// TwinCAT 3 PLC project Conveyor
// ProgramVersion: 3.1.4026.27
// libraries:
//   Tc2_Standard, * (Beckhoff Automation GmbH)
//   Tc2_System, * (Beckhoff Automation GmbH)
//   Tc3_Module, * (Beckhoff Automation GmbH)
// project tree:
//   GVLs/ GVL_IO.TcGVL
//   / PlcTask.TcTTO
//   POUs/ E_ConveyorMode.TcDUT, E_ConveyorState.TcDUT, E_FaultCode.TcDUT, FB_Conveyor.TcPOU, MAIN.TcPOU
// real-time tasks:
//   TASK PlcTask: cycle T#10ms, priority 20, ADS port 350

CONFIGURATION Conveyor
    RESOURCE PLC ON TwinCAT3
        TASK PlcTask(INTERVAL := T#10ms, PRIORITY := 20);
        PROGRAM MAIN WITH PlcTask : MAIN;
    END_RESOURCE
END_CONFIGURATION

// ---- POUs/E_ConveyorMode.TcDUT
{attribute 'qualified_only'}
{attribute 'strict'}
TYPE E_ConveyorMode  :
(
	AUTO,
	MANUAL
);
END_TYPE

// ---- POUs/E_ConveyorState.TcDUT
{attribute 'qualified_only'}
{attribute 'strict'}
TYPE E_ConveyorState :
(
	IDLE,
    RUNNING,
	WAIT_EXIT,
    FAULT
);
END_TYPE

// ---- POUs/E_FaultCode.TcDUT
{attribute 'qualified_only'}
{attribute 'strict'}
TYPE E_FaultCode :
(
	FC_NONE,
	FC_EMERGENCY_STOP,
	FC_EXIT_TIMEOUT
);
END_TYPE

// ---- GVLs/GVL_IO.TcGVL
{attribute 'qualified_only'}
VAR_GLOBAL
	//Input
	StartButton		:	BOOL;
	StopButton		:	BOOL;
	EmergencyStop	:	BOOL;
	Reset			:	BOOL;
	
	SensorEntry		:	BOOL;
	SensorExit		:	BOOL;
	AutoMode		:	BOOL;
	
	
	//Output
	Motor			:	BOOL;
	MotorStopped 	: 	BOOL;
	GreenLamp 		:	BOOL;
	RedLamp 		:	BOOL;
	
	FaultLamp		:	BOOL;
	
	FaultCode 		: 	E_FaultCode;
	
	FaultText : STRING(50) := 'NO FAULT';
	ModeText  : STRING(50) ;
	
	
	Mode : E_ConveyorMode := E_ConveyorMode.AUTO;
	
	
	
	
END_VAR

// ---- POUs/MAIN.TcPOU
PROGRAM MAIN
VAR
	Conveyor		:	FB_Conveyor;
	StartTrigger 	: 	R_TRIG;
	StopTrigger		:	R_TRIG;
	EmergencyOn		:	R_TRIG;
	Reset			:	R_TRIG; 
	
	
	
	
END_VAR

Conveyor(
    Start := GVL_IO.StartButton,
    Stop := GVL_IO.StopButton,
    EmergencyStop := GVL_IO.EmergencyStop,
    Reset := GVL_IO.Reset,
	AutoMode := GVL_IO.AutoMode,
	Mode := GVL_IO.Mode
);

GVL_IO.Motor := Conveyor.Motor;
GVL_IO.MotorStopped := NOT Conveyor.Motor;
GVL_IO.GreenLamp := Conveyor.GreenLamp;
GVL_IO.RedLamp := Conveyor.RedLamp;
GVL_IO.FaultLamp := Conveyor.FaultLamp;
GVL_IO.FaultCode := Conveyor.FaultCode;

GVL_IO.FaultCode := Conveyor.FaultCode;

IF GVL_IO.Mode = E_ConveyorMode.AUTO THEN
	StartTrigger(CLK := GVL_IO.StartButton);
END_IF

StopTrigger(CLK := GVL_IO.StopButton);
EmergencyOn(CLK:= GVL_IO.EmergencyStop);
Reset(CLK:=GVL_IO.Reset);


IF StartTrigger.Q THEN
    GVL_IO.StartButton := FALSE;
END_IF;
IF StopTrigger.Q THEN
	GVL_IO.StopButton := FALSE;
END_IF
IF EmergencyOn.Q THEN
	GVL_IO.EmergencyStop := FALSE;
END_IF
IF Reset.Q THEN
	GVL_IO.Reset := FALSE;
END_IF


CASE GVL_IO.FaultCode OF
    E_FaultCode.FC_NONE:
        GVL_IO.FaultText := 'NO FAULT';

    E_FaultCode.FC_EMERGENCY_STOP:
        GVL_IO.FaultText := 'EMERGENCY STOP';

    E_FaultCode.FC_EXIT_TIMEOUT:
        GVL_IO.FaultText := 'EXIT SENSOR TIMEOUT';
END_CASE

IF GVL_IO.AutoMode THEN
    GVL_IO.Mode := E_ConveyorMode.AUTO;
ELSE
    GVL_IO.Mode := E_ConveyorMode.MANUAL;
END_IF

IF GVL_IO.Mode = E_ConveyorMode.AUTO THEN
	GVL_IO.ModeText := 'AUTO';
ELSIF GVL_IO.Mode = E_ConveyorMode.MANUAL THEN
	GVL_IO.ModeText := 'MANUAL'; 
END_IF

END_PROGRAM

// ---- POUs/FB_Conveyor.TcPOU
FUNCTION_BLOCK FB_Conveyor
VAR_INPUT
	
	Start			:	BOOL;
	Stop			:	BOOL;
	EmergencyStop	:	BOOL;
	Reset			:	BOOL;
	
	AutoMode      	:	BOOL;
	SensorEntry   	: 	BOOL;
    SensorExit    	: 	BOOL;
	
	Mode	:	E_ConveyorMode;
	
END_VAR
VAR_OUTPUT
	
	Motor 		: BOOL;
	GreenLamp 	: BOOL;
	RedLamp 	: BOOL;
	FaultLamp	: BOOL;
	
	FaultCode : E_FaultCode := E_FaultCode.FC_NONE;
	
	
	
END_VAR
VAR
	
   
   
	
	State 	: 	E_ConveyorState ;
	
	
	ModeChanged 	: BOOL;
    PreviousMode 	: E_ConveyorMode;

  
	
	TimerPart		:	TON;
	ExitTrigger		:	R_TRIG;
	EntryTrigger 	: 	R_TRIG;
	Counter 		: 	UDINT := 0;
	
	InterlockOK 	: 	BOOL;
	
	
	
	
	
END_VAR

TimerPart(
    	IN := (Mode = E_ConveyorMode.AUTO)
          	AND 
				(State = E_ConveyorState.WAIT_EXIT),
    	PT := T#10S
	);
ExitTrigger(CLK := SensorExit);	
EntryTrigger(CLK := SensorEntry);
ModeChanged := Mode <> PreviousMode;

IF NOT HandleFaults() THEN
    IF NOT HandleModeChange() THEN
        IF Mode = E_ConveyorMode.AUTO THEN
            RunAuto();

        ELSIF Mode = E_ConveyorMode.MANUAL THEN
            RunManual();
        END_IF
    END_IF
END_IF

UpdateOutputs();

METHOD HandleFaults : BOOL
VAR_INPUT
END_VAR

VAR
END_VAR
HandleFaults := FALSE;

IF EmergencyStop THEN
    State := E_ConveyorState.FAULT;
    FaultCode := E_FaultCode.FC_EMERGENCY_STOP;
    HandleFaults := TRUE;

ELSIF Reset AND State = E_ConveyorState.FAULT THEN
    State := E_ConveyorState.IDLE;
    FaultCode := E_FaultCode.FC_NONE;
    HandleFaults := TRUE;

ELSIF State = E_ConveyorState.FAULT THEN
    HandleFaults := TRUE;
END_IF
END_METHOD

METHOD HandleModeChange : BOOL
VAR_INPUT
END_VAR
HandleModeChange := FALSE;

IF ModeChanged THEN
    IF State <> E_ConveyorState.FAULT THEN
        State := E_ConveyorState.IDLE;
    END_IF

    HandleModeChange := TRUE;
END_IF
END_METHOD

METHOD RunAuto
VAR_INPUT
END_VAR
IF SensorExit THEN
    InterlockOK := FALSE;
ELSE
    InterlockOK := TRUE;
END_IF

CASE State OF

    E_ConveyorState.IDLE:
        IF Start AND InterlockOK THEN
            State := E_ConveyorState.RUNNING;
        END_IF

    E_ConveyorState.RUNNING:
        IF EntryTrigger.Q THEN
            State := E_ConveyorState.WAIT_EXIT;
        ELSIF Stop THEN
            State := E_ConveyorState.IDLE;
        END_IF

    E_ConveyorState.WAIT_EXIT:
        IF TimerPart.Q THEN
            State := E_ConveyorState.FAULT;
            FaultCode := E_FaultCode.FC_EXIT_TIMEOUT;
        ELSIF ExitTrigger.Q THEN
            State := E_ConveyorState.RUNNING;
            Counter := Counter + 1;
        ELSIF Stop THEN
            State := E_ConveyorState.IDLE;
        END_IF

END_CASE
END_METHOD

METHOD RunManual
VAR_INPUT
END_VAR
IF State <> E_ConveyorState.FAULT THEN
    IF Start THEN
        State := E_ConveyorState.RUNNING;
    ELSE
        State := E_ConveyorState.IDLE;
    END_IF
END_IF
END_METHOD

METHOD UpdateOutputs
VAR_INPUT
END_VAR
Motor := (State = E_ConveyorState.RUNNING)
      OR (State = E_ConveyorState.WAIT_EXIT);

GreenLamp := Motor;
RedLamp := State = E_ConveyorState.IDLE;
FaultLamp := State = E_ConveyorState.FAULT;
END_METHOD

END_FUNCTION_BLOCK
